SUBAPPLICATION Uebung_272_AX (* Dialog: Ja/Nein/Abbrechen, Fokus Nein, modal, Ton, nach 10 s RESULT 8 *)
  (* Standard: 61499-2; Description: Copyright (c) 2026 Meisterschulen am Ostbahnhof This program and the accompanying materials are made available under the terms of the Eclipse Public License 2.0 which is available at https://www.eclipse.org/legal/epl-2.0/ SPDX-License-Identifier: EPL-2.0 *)
  (* Version 1.0, 2026-11-17, Franz Höpfinger, Meisterschulen am Ostbahnhof, initial API and implementation and/or initial documentation *)
  PACKAGE Uebungen;
  IMPORT Uebungen::const::UT::Dialog::DefaultPool::OutputNumber_Result;
  IMPORT Uebungen::const::UT::Dialog::DefaultPool::OutputString_Text_Frage;
  IMPORT Uebungen::const::UT::Dialog::DefaultPool::SoftKey_F4;
  IMPORT isobus::UT::dialog::DialogConst::DLG_BTN_YESNOCANCEL;
  IMPORT isobus::UT::dialog::DialogConst::DLG_ICON_QUESTION;
  IMPORT isobus::UT::io::Softkey::SoftKeyActivationCode::SK_RELEASED;
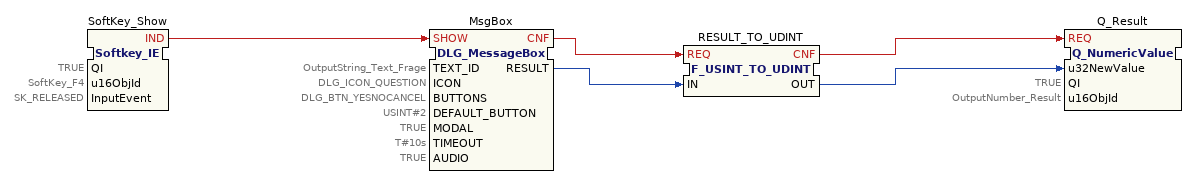
  FBS
    SoftKey_Show : isobus::UT::io::Softkey::Softkey_IE(QI := TRUE, u16ObjId := SoftKey_F4, InputEvent := SK_RELEASED);
    MsgBox : isobus::UT::dialog::DLG_MessageBox(TEXT_ID := OutputString_Text_Frage, ICON := DLG_ICON_QUESTION, BUTTONS := DLG_BTN_YESNOCANCEL, DEFAULT_BUTTON := USINT#2, MODAL := TRUE, TIMEOUT := T#10s, AUDIO := TRUE);
    RESULT_TO_UDINT : iec61131::conversion::F_USINT_TO_UDINT;
    Q_Result : isobus::UT::Q::Q_NumericValue(QI := TRUE, u16ObjId := OutputNumber_Result);
  END_FBS
  EVENT_CONNECTIONS
    SoftKey_Show.IND TO MsgBox.SHOW;
    MsgBox.CNF TO RESULT_TO_UDINT.REQ;
    RESULT_TO_UDINT.CNF TO Q_Result.REQ;
  END_CONNECTIONS
  DATA_CONNECTIONS
    MsgBox.RESULT TO RESULT_TO_UDINT.IN;
    RESULT_TO_UDINT.OUT TO Q_Result.u32NewValue;
  END_CONNECTIONS
END_SUBAPPLICATION
